// TIA Portal V20 export
FUNCTION_BLOCK "OP1"   // FB50, LAD
{ S7_Optimized_Access := 'TRUE' }
// stored: AutoNumber false, MemoryReserve 100, SetENOAutomatically false
   VAR DB_SPECIFIC
      CONTROL_MAN : Struct
         kar_work : Bool;
         kar_home : Bool;
         zarazka_work : Bool;
         zarazka_home : Bool;
         B4 : Bool;
         B5 : Bool;
         B6 : Bool;
         B7 : Bool;
         B8 : Bool;
         B9 : Bool;
         odfuk_1 : Bool;
         odfuk_2 : Bool;
         B12 : Bool;
         B13 : Bool;
         B14 : Bool;
         B15 : Bool;
         B16 : Bool;
         B17 : Bool;
         B18 : Bool;
         B19 : Bool;
         B20 : Bool;
         B21 : Bool;
         B22 : Bool;
         B23 : Bool;
         B24 : Bool;
         B25 : Bool;
         B26 : Bool;
         B27 : Bool;
         B28 : Bool;
         B29 : Bool;
         B30 : Bool;
         B31 : Bool;
      END_STRUCT;
      CONTROL_AUTOMAT : Struct
         KAR_WORK : Bool;
         KAR_HOME : Bool;
         ZARAZKA_WORK : Bool;
         ZARAZKA_HOME : Bool;
         B4 : Bool;
         B5 : Bool;
         B6 : Bool;
         B7 : Bool;
         B8 : Bool;
         B9 : Bool;
         odfuk_1 : Bool;
         odfuk_2 : Bool;
         B12 : Bool;
         B13 : Bool;
         B14 : Bool;
         B15 : Bool;
         B16 : Bool;
         B17 : Bool;
         B18 : Bool;
         B19 : Bool;
         B20 : Bool;
         B21 : Bool;
         B22 : Bool;
         B23 : Bool;
         B24 : Bool;
         B25 : Bool;
         B26 : Bool;
         B27 : Bool;
         B28 : Bool;
         B29 : Bool;
         B30 : Bool;
         B31 : Bool;
      END_STRUCT;
      SENSORS : Struct
         prechod_1 : Bool;
         prechod_1_neg : Bool;
         kontrola : Bool;
         kontrola_neg : Bool;
         prechod_2 : Bool;
         Prechod_2_neg : Bool;
         Pozice_vyrazovace : Bool;
         Pozice_vyrazovace_neg : Bool;
         Pozice_pistu : Bool;   // KARUSEL JE NATOČEN PŘÍPRAVKEM A K BRÁNĚ
         Pozice_pistu_neg : Bool;
         s10 : Bool;
         s11 : Bool;
         s12 : Bool;
         s13 : Bool;
         s14 : Bool;
         s15 : Bool;
         s16 : Bool;
         s17 : Bool;
         s18 : Bool;
         s19 : Bool;
         s20 : Bool;
         s21 : Bool;
         s22 : Bool;
         s23 : Bool;
         s24 : Bool;
         s25 : Bool;
         s26 : Bool;
         s27 : Bool;
         s28 : Bool;
         s29 : Bool;
         s30 : Bool;
         s31 : Bool;
      END_STRUCT;
      SENSORS_1 : Struct
         S0 : Bool;
         S1 : Bool;
         S2 : Bool;
         S3 : Bool;
         S4 : Bool;
         S5 : Bool;
         S6 : Bool;
         S7 : Bool;
         S8 : Bool;
         S9 : Bool;
         SESTAVA_NENI_OTOCENA : Bool;
         SESTAVA_JE_OTOCENA : Bool;
         S12 : Bool;
         S13 : Bool;
         S14 : Bool;
         S15 : Bool;
         S16 : Bool;
         S17 : Bool;
         S18 : Bool;
         S19 : Bool;
         S20 : Bool;
         S21 : Bool;
         S22 : Bool;
         S23 : Bool;
         S24 : Bool;
         S25 : Bool;
         S26 : Bool;
         S27 : Bool;
         S28 : Bool;
         S29 : Bool;
         S30 : Bool;
         l_3_neg : Bool;
      END_STRUCT;
   END_VAR
   VAR
      S_0 : "SENSOR";
      S_1 : "SENSOR";
      S_2 { S7_SetPoint := 'True'} : "SENSOR";
      S_3 { S7_SetPoint := 'True'} : "SENSOR";
      S_4 { S7_SetPoint := 'True'} : "SENSOR";
      S_5 { S7_SetPoint := 'True'} : "SENSOR";
      S_6 { S7_SetPoint := 'True'} : "SENSOR";
      M_karusel : "MOTOR_CONTROL_BLOCK";
      M_zarazka { S7_SetPoint := 'True'} : "MOTOR_CONTROL_BLOCK";
      M_CLONA { S7_SetPoint := 'True'} : "MOTOR_CONTROL_BLOCK";
   END_VAR
   VAR DB_SPECIFIC
      SQCR { S7_SetPoint := 'True'} : Int;
   END_VAR
   VAR
      hmi_sqcr : Int;
   END_VAR
   VAR DB_SPECIFIC
      TRIG : Struct
         inicial_ok_op : Bool;
         DSSAD : Bool;
         INICIALIZACE_PROBEHLA : Bool;
         trig_dil : Bool;
         p_trig_control_tcon : Bool;
         T6 : Bool;
         SPUST_OP_4 : Bool;
         vlez_do_zavory_pri_rotaci : Bool;
         START_INICIAL_OP2 : Bool;
         START_INICIAL_OP3 : Bool;
         spust_odsavani : Bool;
         VYPRAZNI_OK_OP_2_A : Bool;
         VYPRAZNI_NOK_OP_2_A : Bool;
         VYPRAZDNI_OK_OP_3_B : Bool;
         VYPRAZDNI_NOK_OP_3_B : Bool;
         RESET_NCODER : Bool;
         op_1_ready : Bool;
      END_STRUCT;
      MEMOR : Struct
         n_trig_vypnuti : Bool;
         M1 : Bool;
         M2 : Bool;
         M3 : Bool;
         M4 : Bool;
         p_trig_odavacka : Bool;
         M6 : Bool;
         M7 : Bool;
         M8 : Bool;
         M9 : Bool;
         M10 : Bool;
         M11 : Bool;
         RESET_ERROR : Bool;
         vyrazeni_pamet : Bool;
         M14 : Bool;
         M15 : Bool;
         SETOVANI_START : Bool;
         M17 : Bool;
         p_trig_pamet_1 : Bool;
         p_trig_pamet_2 : Bool;
         p_trig_pamet_3 : Bool;
         p_trig_pamet_4 : Bool;
         p_trig_pamet_5 : Bool;
         p_trig_pamet_6 : Bool;
         p_trig_pamet_7 : Bool;
         p_trig_pamet_8 : Bool;
         p_trig_pamet_9 : Bool;
         p_trig_pamet_10 : Bool;
         p_trig_vyrad : Bool;
         p_Trig_cisteni_pozice : Bool;
         p_trig_citac : Bool;
         N_TRIG_SAFETY : Bool;
         P_TRIG_RESET_POZICE : Bool;
         M33 : Bool;
         start_caklu : Bool;
         M35 : Bool;
         M36 : Bool;
         M37 : Bool;
         M38 : Bool;
         M39 : Bool;
         ALARM_GLOBAL : Bool;
         M41 : Bool;
         M42 : Bool;
         M43 : Bool;
         M44 : Bool;
         M45 : Bool;
         M46 : Bool;
         M47 : Bool;
         M48 : Bool;
         M49 : Bool;
         wrong_p_trig : Bool;
         alarm_p_trig : Bool;
         M52 : Bool;
         M53 : Bool;
         M54 : Bool;
         M55 : Bool;
         M56 : Bool;
         M57 : Bool;
         M58 : Bool;
         M59 : Bool;
         M60 : Bool;
         M61 : Bool;
         M62 : Bool;
         M63 : Bool;
      END_STRUCT;
      "TIMER" : Struct
         TIMER_0 : IEC_TIMER;
         TIMER_VACUUM_CLEANER : IEC_TIMER;
         TIMER_DELAY_RESET_EXECUTE : IEC_TIMER;
         TIMER_3 : IEC_TIMER;
         TIMER_4 : IEC_TIMER;
         air : IEC_TIMER;
         TIMER_6 : IEC_TIMER;
         TIMER_7 : IEC_TIMER;
      END_STRUCT;
      HMI : Struct
         povoleni_volby_receptu : Bool;
         "svetlo_on/off" : Bool;
         ALARM_VIDITELNOST : Bool;
         hmi_3 : Bool;
         hmi_4 : Bool;
         reset_fronty : Bool;
         hmi_6 : Bool;
         hmi_7 : Bool;
         hmi_8 : Bool;
         hmi_9 : Bool;
         hmi_10 : Bool;
         hmi_11 : Bool;
         hmi_12 : Bool;
         hmi_13 : Bool;
         hmi_14 : Bool;
         hmi_15 : Bool;
      END_STRUCT;
   END_VAR
   VAR
      STRING_0 : String[1];
      array_chyb_ctec : Array[1..16] of Bool;
      zpracovani_dat { ExternalAccessible := 'False'; ExternalVisible := 'False'; ExternalWritable := 'False'} : Array[1..1] of Struct
         prenaseny_text : String[100];
         balik_den : Int;
         vyrazeni : Bool;
      END_STRUCT;
   END_VAR
   VAR DB_SPECIFIC
      aktual_kusy : Int;
   END_VAR
   VAR
      i : Int;
      q : Int;
      pocet_znaku_string_kamera : Int;
      ocekavany_text : String[100];
      format_etiketa_ok : Bool;
      Kamera : Struct
         s2_pamet : Bool;
         s2_nabeh : Bool;
         sber_aktivni : Bool;
         prijato_etiketa : Bool;
         prijato_folie_l : Bool;
         prijato_folie_p : Bool;
         ok_etiketa : Bool;
         ok_folie_l : Bool;
         ok_folie_p : Bool;
         vyradit : Bool;
         fronta_plna : Bool;   // alarm
         bypass_ocr : Bool := True;   // dočasně, dokud není doladěné OCR
         last_id_etiketa : Word;
         last_id_folie_l : Word;
         last_id_folie_p : Word;
         balik_den : Int;
         idx : Int;
         pocet : Int;
         text_etiketa : String[100];
         timeout_sberu : Time :=  T#1S;
         kontrola_tridirny : Bool := true;   // HMI: kontrola kódu třídírny zapnuta
         tridirna_ok : Bool;   // výsledek kontroly posledního plata (pro online diagnostiku)
      END_STRUCT;
      Vyrazeni : Struct
         s4_pamet : Bool;
         s4_nabeh : Bool;
         aktivni : Bool;
         vyradit : Bool;
         chyba_bez_dat : Bool;   // alarm: plato u vyřazovače bez záznamu
         chyba_pist : Bool;   // alarm: píst nevyjel / nebyl v home
         max_puls : Time := T#200MS;
         vyrazovac_pripojen : Bool := true;   // TRUE až bude signál od dodavatele
         alarm_nok_balik : Bool;   // NOK plato prošlo bez vyřazení
         posledni_nok_balik : Int;   // číslo plata pro obsluhu / HMI
         posledni_nok_text : String[100];   // co přečetla kamera
         pocet_nok : DInt;   // počítadlo NOK plat
         pocet_bez_dat : DInt;
         majak_tp : TP_TIME;   // prodlouzeni blikani majaku pri vzrazenii
         majak { S7_SetPoint := 'True'} : Bool;
      END_STRUCT;
      Kam_Etiketa_Job : Struct
         krok : Int;   // 0 klid, 10 odeslat, 20 čekat, 30 ukončit handshake
         pozadovany : Int;   // job z receptury (PRG_CAM_etiketa)
         odesli_pamet : Bool;   // hrana ODESLI_dATA
         aktivni : Bool;   // probíhá načítání jobu → blokovat triggery
         chyba : Bool;   // alarm: job se nepodařilo načíst
         chyba_kod : Word;   // CommandResultCode při chybě
         nesouhlasi : Bool;   // alarm: job v kameře ≠ job z receptury
         timeout : Time := T#10S;   // max. doba načítání jobu
      END_STRUCT;
      Test_tp_ka12 : TP_TIME;
   END_VAR
   VAR_TEMP
      DATA : Array[0..255] of Char;
      ARRAY_NULL : Array[1..8] of Bool;
      array_null_fronta : Array[1..1] of Struct
         prenaseny_text : String[100];
         balik_den : Int;
         vyrazeni : Bool;
      END_STRUCT;
      "char" : Array[0..0] of Char;
      "string" : String;
      cas : DTL;
      ret : Int;
   END_VAR
   VAR CONSTANT
      STEP_0 : Int := 0;
      step_2 : Int := 2;
      STEP_4 : Int := 4;
      STEP_5_HOME : Int := 5;
      STEP_7 : Int := 7;
      STEP_10 : Int := 10;
      STEP_15 : Int := 15;
      STEP_20 : Int := 20;
      STEP_23 : Int := 23;
      STEP_25 : Int := 25;
      STEP_27 : Int := 27;
      STEP_30 : Int := 30;
      STEP_35 : Int := 35;
      STEP_37 : Int := 37;
      STEP_40 : Int := 40;
      STEP_45 : Int := 45;
      STEP_50 : Int := 50;
      STEP_55 : Int := 55;
      STEP_60 : Int := 60;
      STEP_65 : Int := 65;
      STEP_70 : Int := 70;
      STEP_75 : Int := 75;
      STEP_80 : Int := 80;
      STEP_83 : Int := 83;
      STEP_85 : Int := 85;
      STEP_90 : Int := 90;
      STEP_95 : Int := 95;
      STEP_100 : Int := 100;
      STEP_105 : Int := 105;
      STEP_110 : Int := 110;
      STEP_113 : Int := 113;
      STEP_115 : Int := 115;
      STEP_120 : Int := 120;
      STEP_125 : Int := 125;
      STEP_130 : Int := 130;
      STEP_135 : Int := 135;
      STEP_140 : Int := 140;
      STEP_145 : Int := 145;
      STEP_150 : Int := 150;
      STEP_155 : Int := 155;
      STEP_1000 : Int := 1000;
      STEP_1001 : Int := 1001;
      STEP_1002 : Int := 1002;
      STEP_1003 : Int := 1003;
      STEP_1004 : Int := 1004;
      STEP_1005 : Int := 1005;
      STEP_1010 : Int := 1010;
      STEP_1015 : Int := 1015;
      STEP_1020 : Int := 1020;
      STEP_1025 : Int := 1025;
      STEP_3000 : Int := 3000;
      STEP_3005 : Int := 3005;
      STEP_3010 : Int := 3010;
      STEP_3015 : Int := 3015;
      STEP_3020 : Int := 3020;
      STEP_2000 : Int := 2000;
      string_null : String;
      char_null : Char;
      text_kartacek : String := 'Kartacek';
      string_kar_A : String := 'A';
      string_kar_B : String := 'B';
      KOD_TRIDIRNY : String := 'CZ32880102';
   END_VAR
   VAR_TEMP   // added for the SCL form of the ladder/FBD networks
      _w1 : Bool;
      _w2 : Bool;
      _w3 : Bool;
   END_VAR
BEGIN

REGION Network 1: manuali ovladani reset
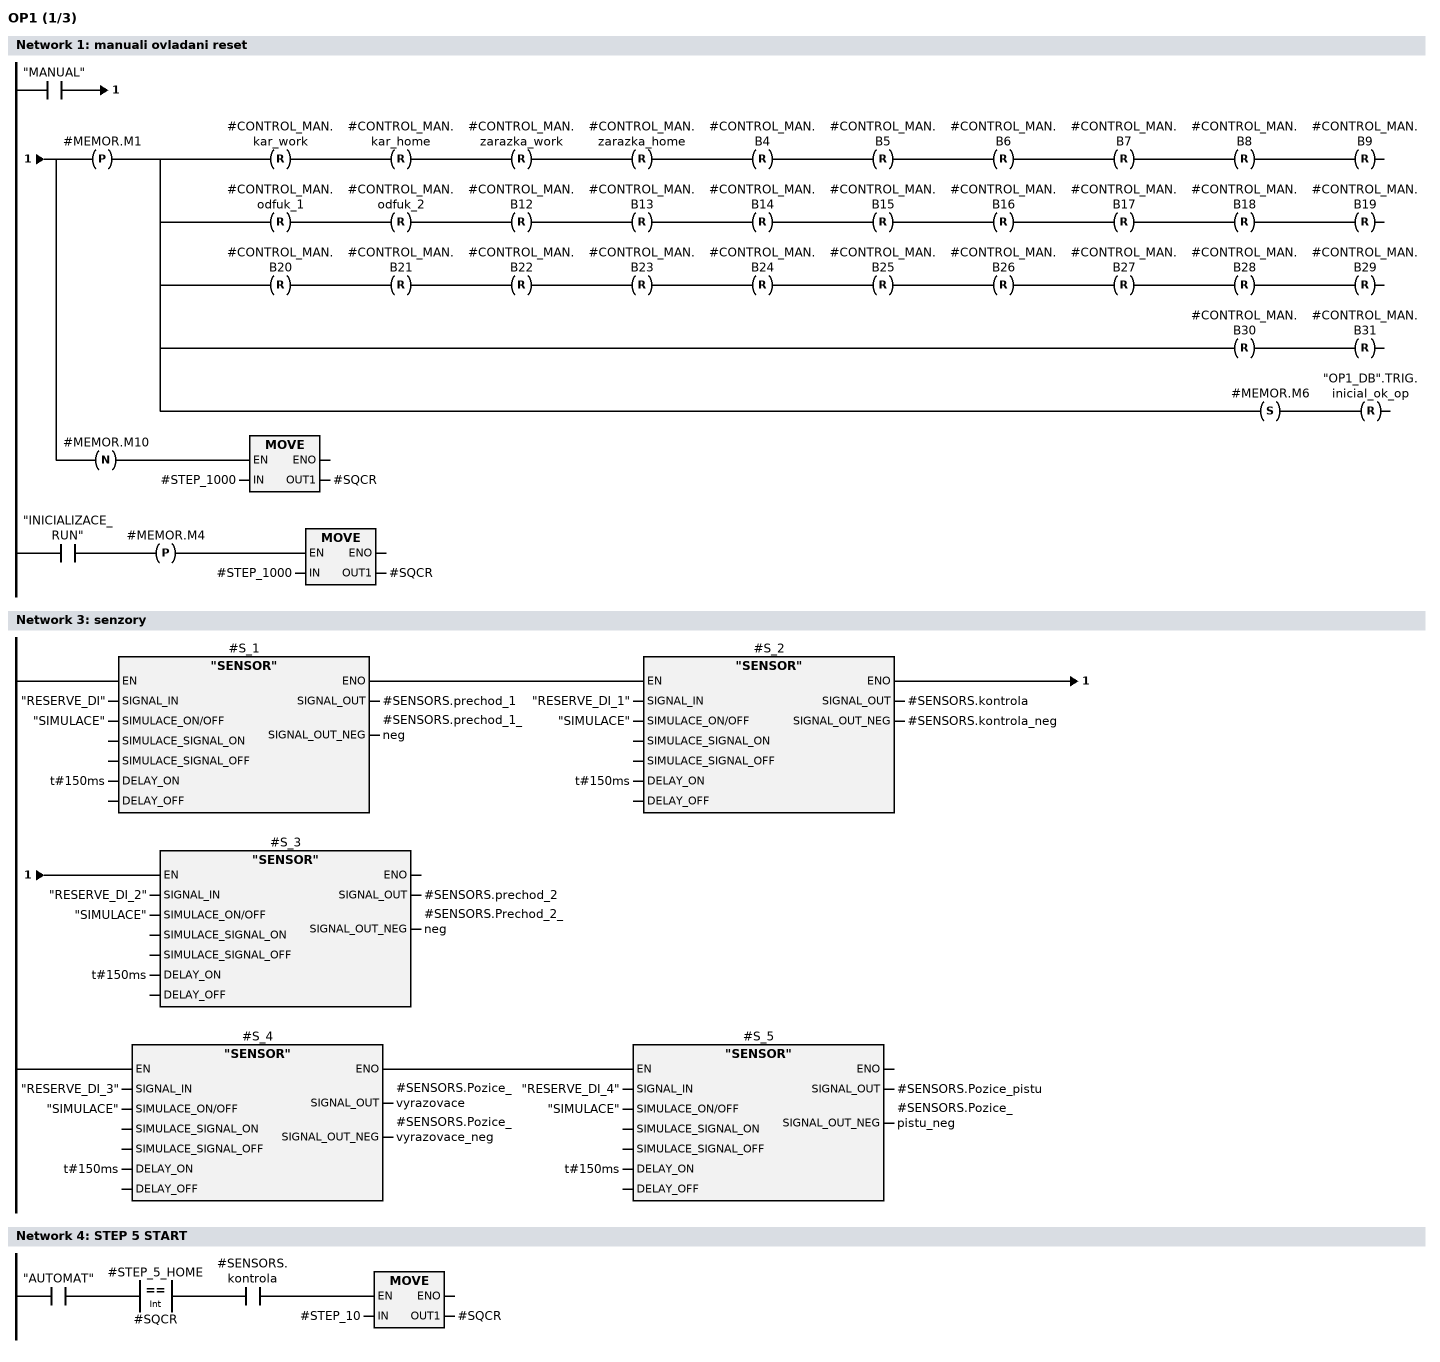
   RUNG wire#powerrail
      Contact( "MANUAL" )
      wire#w1
      P_Trig( #MEMOR.M1 )
      wire#w2
      R_Coil( #CONTROL_MAN.kar_work )
      R_Coil( #CONTROL_MAN.kar_home )
      R_Coil( #CONTROL_MAN.zarazka_work )
      R_Coil( #CONTROL_MAN.zarazka_home )
      R_Coil( #CONTROL_MAN.B4 )
      R_Coil( #CONTROL_MAN.B5 )
      R_Coil( #CONTROL_MAN.B6 )
      R_Coil( #CONTROL_MAN.B7 )
      R_Coil( #CONTROL_MAN.B8 )
      R_Coil( #CONTROL_MAN.B9 )
   END_RUNG
   RUNG wire#w2
      R_Coil( #CONTROL_MAN.odfuk_1 )
      R_Coil( #CONTROL_MAN.odfuk_2 )
      R_Coil( #CONTROL_MAN.B12 )
      R_Coil( #CONTROL_MAN.B13 )
      R_Coil( #CONTROL_MAN.B14 )
      R_Coil( #CONTROL_MAN.B15 )
      R_Coil( #CONTROL_MAN.B16 )
      R_Coil( #CONTROL_MAN.B17 )
      R_Coil( #CONTROL_MAN.B18 )
      R_Coil( #CONTROL_MAN.B19 )
   END_RUNG
   RUNG wire#w2
      R_Coil( #CONTROL_MAN.B20 )
      R_Coil( #CONTROL_MAN.B21 )
      R_Coil( #CONTROL_MAN.B22 )
      R_Coil( #CONTROL_MAN.B23 )
      R_Coil( #CONTROL_MAN.B24 )
      R_Coil( #CONTROL_MAN.B25 )
      R_Coil( #CONTROL_MAN.B26 )
      R_Coil( #CONTROL_MAN.B27 )
      R_Coil( #CONTROL_MAN.B28 )
      R_Coil( #CONTROL_MAN.B29 )
   END_RUNG
   RUNG wire#w2
      R_Coil( #CONTROL_MAN.B30 )
      R_Coil( #CONTROL_MAN.B31 )
   END_RUNG
   RUNG wire#w2
      S_Coil( #MEMOR.M6 )
      R_Coil( "OP1_DB".TRIG.inicial_ok_op )
   END_RUNG
   RUNG wire#w1
      N_Trig( #MEMOR.M10 )
      Move(in := #STEP_1000, out1 => #SQCR)
   END_RUNG
   RUNG wire#powerrail
      Contact( "INICIALIZACE_RUN" )
      P_Trig( #MEMOR.M4 )
      Move(in := #STEP_1000, out1 => #SQCR)
   END_RUNG
   // the same network as SCL:
   #_w1 := "MANUAL" AND NOT #MEMOR.M1;   // rising edge
   #MEMOR.M1 := "MANUAL";
   IF #_w1 THEN
       #CONTROL_MAN.kar_work := FALSE;
       #CONTROL_MAN.kar_home := FALSE;
       #CONTROL_MAN.zarazka_work := FALSE;
       #CONTROL_MAN.zarazka_home := FALSE;
       #CONTROL_MAN.B4 := FALSE;
       #CONTROL_MAN.B5 := FALSE;
       #CONTROL_MAN.B6 := FALSE;
       #CONTROL_MAN.B7 := FALSE;
       #CONTROL_MAN.B8 := FALSE;
       #CONTROL_MAN.B9 := FALSE;
       #CONTROL_MAN.odfuk_1 := FALSE;
       #CONTROL_MAN.odfuk_2 := FALSE;
       #CONTROL_MAN.B12 := FALSE;
       #CONTROL_MAN.B13 := FALSE;
       #CONTROL_MAN.B14 := FALSE;
       #CONTROL_MAN.B15 := FALSE;
       #CONTROL_MAN.B16 := FALSE;
       #CONTROL_MAN.B17 := FALSE;
       #CONTROL_MAN.B18 := FALSE;
       #CONTROL_MAN.B19 := FALSE;
       #CONTROL_MAN.B20 := FALSE;
       #CONTROL_MAN.B21 := FALSE;
       #CONTROL_MAN.B22 := FALSE;
       #CONTROL_MAN.B23 := FALSE;
       #CONTROL_MAN.B24 := FALSE;
       #CONTROL_MAN.B25 := FALSE;
       #CONTROL_MAN.B26 := FALSE;
       #CONTROL_MAN.B27 := FALSE;
       #CONTROL_MAN.B28 := FALSE;
       #CONTROL_MAN.B29 := FALSE;
       #CONTROL_MAN.B30 := FALSE;
       #CONTROL_MAN.B31 := FALSE;
       #MEMOR.M6 := TRUE;
       "OP1_DB".TRIG.inicial_ok_op := FALSE;
   END_IF;
   #_w2 := NOT "MANUAL" AND #MEMOR.M10;   // falling edge
   #MEMOR.M10 := "MANUAL";
   IF #_w2 THEN #SQCR := #STEP_1000; END_IF;
   #_w3 := "INICIALIZACE_RUN" AND NOT #MEMOR.M4;   // rising edge
   #MEMOR.M4 := "INICIALIZACE_RUN";
   IF #_w3 THEN #SQCR := #STEP_1000; END_IF;
END_REGION

REGION Network 2: alarmy
END_REGION

REGION Network 3: senzory
   RUNG wire#powerrail
      #S_1(SIGNAL_IN := "RESERVE_DI", "SIMULACE_ON/OFF" := "SIMULACE", SIMULACE_SIGNAL_ON :=, SIMULACE_SIGNAL_OFF :=, DELAY_ON := t#150ms, DELAY_OFF :=, SIGNAL_OUT => #SENSORS.prechod_1, SIGNAL_OUT_NEG => #SENSORS.prechod_1_neg)
      #S_2(SIGNAL_IN := "RESERVE_DI_1", "SIMULACE_ON/OFF" := "SIMULACE", SIMULACE_SIGNAL_ON :=, SIMULACE_SIGNAL_OFF :=, DELAY_ON := t#150ms, DELAY_OFF :=, SIGNAL_OUT => #SENSORS.kontrola, SIGNAL_OUT_NEG => #SENSORS.kontrola_neg)
      #S_3(SIGNAL_IN := "RESERVE_DI_2", "SIMULACE_ON/OFF" := "SIMULACE", SIMULACE_SIGNAL_ON :=, SIMULACE_SIGNAL_OFF :=, DELAY_ON := t#150ms, DELAY_OFF :=, SIGNAL_OUT => #SENSORS.prechod_2, SIGNAL_OUT_NEG => #SENSORS.Prechod_2_neg)
   END_RUNG
   RUNG wire#powerrail
      #S_4(SIGNAL_IN := "RESERVE_DI_3", "SIMULACE_ON/OFF" := "SIMULACE", SIMULACE_SIGNAL_ON :=, SIMULACE_SIGNAL_OFF :=, DELAY_ON := t#150ms, DELAY_OFF :=, SIGNAL_OUT => #SENSORS.Pozice_vyrazovace, SIGNAL_OUT_NEG => #SENSORS.Pozice_vyrazovace_neg)
      #S_5(SIGNAL_IN := "RESERVE_DI_4", "SIMULACE_ON/OFF" := "SIMULACE", SIMULACE_SIGNAL_ON :=, SIMULACE_SIGNAL_OFF :=, DELAY_ON := t#150ms, DELAY_OFF :=, SIGNAL_OUT => #SENSORS.Pozice_pistu, SIGNAL_OUT_NEG => #SENSORS.Pozice_pistu_neg)
   END_RUNG
   // the same network as SCL:
   #S_1(SIGNAL_IN := "RESERVE_DI",   // "SENSOR"
        "SIMULACE_ON/OFF" := "SIMULACE",
        DELAY_ON := t#150ms,
        SIGNAL_OUT => #SENSORS.prechod_1,
        SIGNAL_OUT_NEG => #SENSORS.prechod_1_neg,
        ENO => #_w1);
   #S_2(EN := #_w1,   // "SENSOR"
        SIGNAL_IN := "RESERVE_DI_1",
        "SIMULACE_ON/OFF" := "SIMULACE",
        DELAY_ON := t#150ms,
        SIGNAL_OUT => #SENSORS.kontrola,
        SIGNAL_OUT_NEG => #SENSORS.kontrola_neg,
        ENO => #_w2);
   IF #_w2 THEN
       #S_3(SIGNAL_IN := "RESERVE_DI_2",   // "SENSOR"
            "SIMULACE_ON/OFF" := "SIMULACE",
            DELAY_ON := t#150ms,
            SIGNAL_OUT => #SENSORS.prechod_2,
            SIGNAL_OUT_NEG => #SENSORS.Prechod_2_neg);
   END_IF;
   #S_4(SIGNAL_IN := "RESERVE_DI_3",   // "SENSOR"
        "SIMULACE_ON/OFF" := "SIMULACE",
        DELAY_ON := t#150ms,
        SIGNAL_OUT => #SENSORS.Pozice_vyrazovace,
        SIGNAL_OUT_NEG => #SENSORS.Pozice_vyrazovace_neg,
        ENO => #_w3);
   IF #_w3 THEN
       #S_5(SIGNAL_IN := "RESERVE_DI_4",   // "SENSOR"
            "SIMULACE_ON/OFF" := "SIMULACE",
            DELAY_ON := t#150ms,
            SIGNAL_OUT => #SENSORS.Pozice_pistu,
            SIGNAL_OUT_NEG => #SENSORS.Pozice_pistu_neg);
   END_IF;
END_REGION

REGION Network 4: STEP 5 START
   RUNG wire#powerrail
      Contact( "AUTOMAT" )
      { S7_Templates := "SrcType := Int" } EQ_Contact(in1 := #STEP_5_HOME, in2 := #SQCR)
      Contact( #SENSORS.kontrola )
      Move(in := #STEP_10, out1 => #SQCR)
   END_RUNG
   // the same network as SCL:
   IF "AUTOMAT" AND (#STEP_5_HOME = #SQCR) AND #SENSORS.kontrola THEN #SQCR := #STEP_10; END_IF;
END_REGION

REGION Network 5: STEP 10
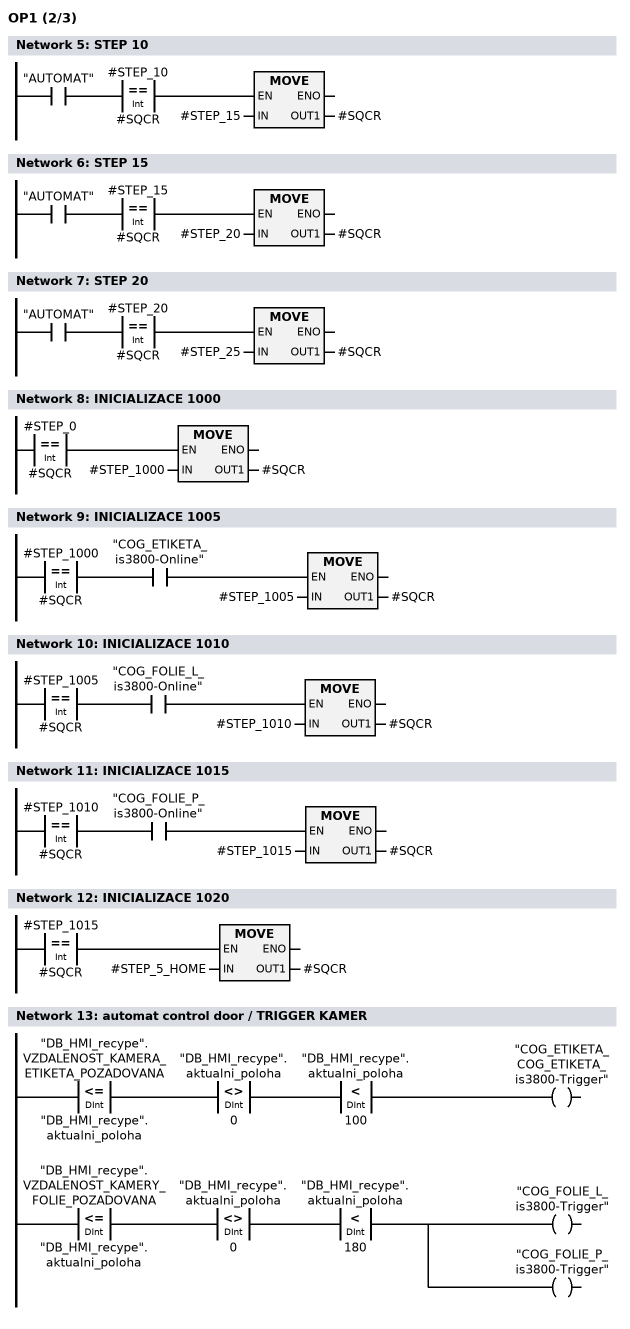
   RUNG wire#powerrail
      Contact( "AUTOMAT" )
      { S7_Templates := "SrcType := Int" } EQ_Contact(in1 := #STEP_10, in2 := #SQCR)
      Move(in := #STEP_15, out1 => #SQCR)
   END_RUNG
   // the same network as SCL:
   IF "AUTOMAT" AND (#STEP_10 = #SQCR) THEN #SQCR := #STEP_15; END_IF;
END_REGION

REGION Network 6: STEP 15
   RUNG wire#powerrail
      Contact( "AUTOMAT" )
      { S7_Templates := "SrcType := Int" } EQ_Contact(in1 := #STEP_15, in2 := #SQCR)
      Move(in := #STEP_20, out1 => #SQCR)
   END_RUNG
   // the same network as SCL:
   IF "AUTOMAT" AND (#STEP_15 = #SQCR) THEN #SQCR := #STEP_20; END_IF;
END_REGION

REGION Network 7: STEP 20
   RUNG wire#powerrail
      Contact( "AUTOMAT" )
      { S7_Templates := "SrcType := Int" } EQ_Contact(in1 := #STEP_20, in2 := #SQCR)
      Move(in := #STEP_25, out1 => #SQCR)
   END_RUNG
   // the same network as SCL:
   IF "AUTOMAT" AND (#STEP_20 = #SQCR) THEN #SQCR := #STEP_25; END_IF;
END_REGION

REGION Network 8: INICIALIZACE 1000
   RUNG wire#powerrail
      { S7_Templates := "SrcType := Int" } EQ_Contact(in1 := #STEP_0, in2 := #SQCR)
      Move(in := #STEP_1000, out1 => #SQCR)
   END_RUNG
   // the same network as SCL:
   IF #STEP_0 = #SQCR THEN #SQCR := #STEP_1000; END_IF;
END_REGION

REGION Network 9: INICIALIZACE 1005
   RUNG wire#powerrail
      { S7_Templates := "SrcType := Int" } EQ_Contact(in1 := #STEP_1000, in2 := #SQCR)
      Contact( "COG_ETIKETA_is3800-Online" )
      Move(in := #STEP_1005, out1 => #SQCR)
   END_RUNG
   // the same network as SCL:
   IF (#STEP_1000 = #SQCR) AND "COG_ETIKETA_is3800-Online" THEN #SQCR := #STEP_1005; END_IF;
END_REGION

REGION Network 10: INICIALIZACE 1010
   RUNG wire#powerrail
      { S7_Templates := "SrcType := Int" } EQ_Contact(in1 := #STEP_1005, in2 := #SQCR)
      Contact( "COG_FOLIE_L_is3800-Online" )
      Move(in := #STEP_1010, out1 => #SQCR)
   END_RUNG
   // the same network as SCL:
   IF (#STEP_1005 = #SQCR) AND "COG_FOLIE_L_is3800-Online" THEN #SQCR := #STEP_1010; END_IF;
END_REGION

REGION Network 11: INICIALIZACE 1015
   RUNG wire#powerrail
      { S7_Templates := "SrcType := Int" } EQ_Contact(in1 := #STEP_1010, in2 := #SQCR)
      Contact( "COG_FOLIE_P_is3800-Online" )
      Move(in := #STEP_1015, out1 => #SQCR)
   END_RUNG
   // the same network as SCL:
   IF (#STEP_1010 = #SQCR) AND "COG_FOLIE_P_is3800-Online" THEN #SQCR := #STEP_1015; END_IF;
END_REGION

REGION Network 12: INICIALIZACE 1020
   RUNG wire#powerrail
      { S7_Templates := "SrcType := Int" } EQ_Contact(in1 := #STEP_1015, in2 := #SQCR)
      Move(in := #STEP_5_HOME, out1 => #SQCR)
   END_RUNG
   // the same network as SCL:
   IF #STEP_1015 = #SQCR THEN #SQCR := #STEP_5_HOME; END_IF;
END_REGION

REGION Network 13: automat control door / TRIGGER KAMER
   RUNG wire#powerrail
      { S7_Templates := "SrcType := DInt" } LE_Contact(in1 := "DB_HMI_recype".VZDALENOST_KAMERA_ETIKETA_POZADOVANA, in2 := "DB_HMI_recype".aktualni_poloha)
      { S7_Templates := "SrcType := DInt" } NE_Contact(in1 := "DB_HMI_recype".aktualni_poloha, in2 := 0)
      { S7_Templates := "SrcType := DInt" } LT_Contact(in1 := "DB_HMI_recype".aktualni_poloha, in2 := 100)
      Coil( "COG_ETIKETA_COG_ETIKETA_is3800-Trigger" )
   END_RUNG
   RUNG wire#powerrail
      { S7_Templates := "SrcType := DInt" } LE_Contact(in1 := "DB_HMI_recype".VZDALENOST_KAMERY_FOLIE_POZADOVANA, in2 := "DB_HMI_recype".aktualni_poloha)
      { S7_Templates := "SrcType := DInt" } NE_Contact(in1 := "DB_HMI_recype".aktualni_poloha, in2 := 0)
      { S7_Templates := "SrcType := DInt" } LT_Contact(in1 := "DB_HMI_recype".aktualni_poloha, in2 := 180)
      wire#w1
      Coil( "COG_FOLIE_L_is3800-Trigger" )
   END_RUNG
   RUNG wire#w1
      Coil( "COG_FOLIE_P_is3800-Trigger" )
   END_RUNG
   // the same network as SCL:
   "COG_ETIKETA_COG_ETIKETA_is3800-Trigger" := ("DB_HMI_recype".VZDALENOST_KAMERA_ETIKETA_POZADOVANA <= "DB_HMI_recype".aktualni_poloha) AND ("DB_HMI_recype".aktualni_poloha <> 0) AND ("DB_HMI_recype".aktualni_poloha < 100);
   "COG_FOLIE_L_is3800-Trigger" := ("DB_HMI_recype".VZDALENOST_KAMERY_FOLIE_POZADOVANA <= "DB_HMI_recype".aktualni_poloha) AND ("DB_HMI_recype".aktualni_poloha <> 0) AND ("DB_HMI_recype".aktualni_poloha < 180);
   "COG_FOLIE_P_is3800-Trigger" := "COG_FOLIE_L_is3800-Trigger";
END_REGION

REGION Network 14: TRIGGER SVETEL
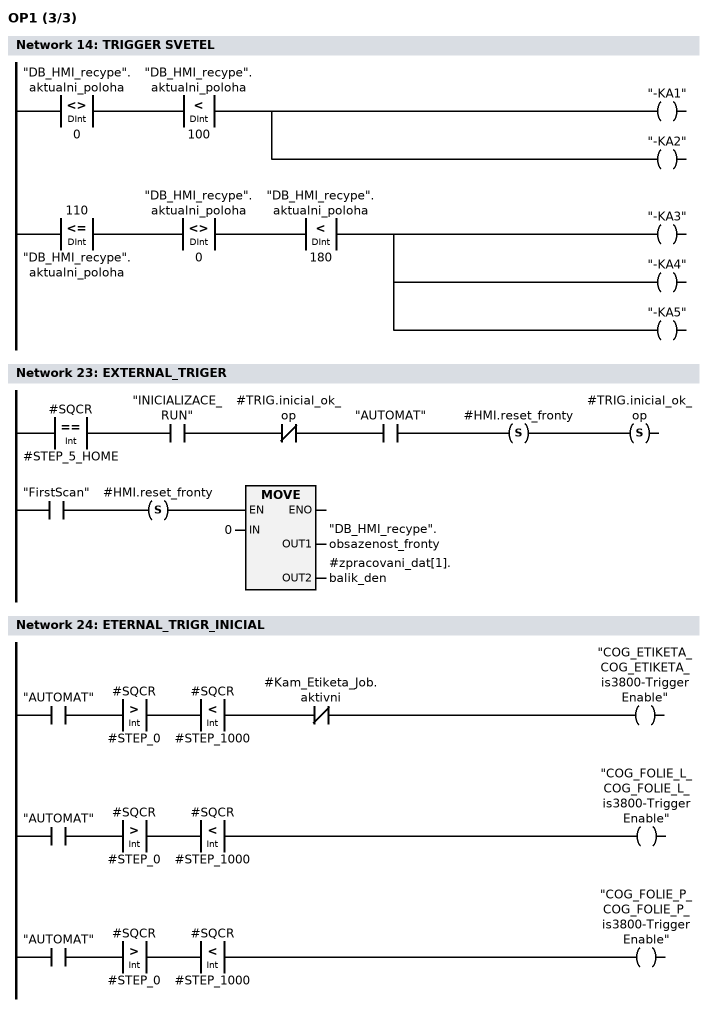
   RUNG wire#powerrail
      { S7_Templates := "SrcType := DInt" } NE_Contact(in1 := "DB_HMI_recype".aktualni_poloha, in2 := 0)
      { S7_Templates := "SrcType := DInt" } LT_Contact(in1 := "DB_HMI_recype".aktualni_poloha, in2 := 100)
      wire#w1
      Coil( "-KA1" )
   END_RUNG
   RUNG wire#w1
      Coil( "-KA2" )
   END_RUNG
   RUNG wire#powerrail
      { S7_Templates := "SrcType := DInt" } LE_Contact(in1 := 110, in2 := "DB_HMI_recype".aktualni_poloha)
      { S7_Templates := "SrcType := DInt" } NE_Contact(in1 := "DB_HMI_recype".aktualni_poloha, in2 := 0)
      { S7_Templates := "SrcType := DInt" } LT_Contact(in1 := "DB_HMI_recype".aktualni_poloha, in2 := 180)
      wire#w2
      Coil( "-KA3" )
   END_RUNG
   RUNG wire#w2
      Coil( "-KA4" )
   END_RUNG
   RUNG wire#w2
      Coil( "-KA5" )
   END_RUNG
   // the same network as SCL:
   "-KA1" := ("DB_HMI_recype".aktualni_poloha <> 0) AND ("DB_HMI_recype".aktualni_poloha < 100);
   "-KA2" := "-KA1";
   "-KA3" := (110 <= "DB_HMI_recype".aktualni_poloha) AND ("DB_HMI_recype".aktualni_poloha <> 0) AND ("DB_HMI_recype".aktualni_poloha < 180);
   "-KA4" := "-KA3";
   "-KA5" := "-KA3";
END_REGION

REGION Network 15 (SCL): TRIGGER MANUAL
   "iDB_CamManual"(xManEtiketa:="DB_Manual".xManEtiketa,
                   xManFolie:="DB_Manual".xManFolie);
END_REGION

REGION Network 16 (SCL): automat control data
   // Smyčka projde 104 bajtů (od 0 do 103)
   FOR #i := 0 TO 103 DO
       // PEEK čte přímo z paměti vstupů (16#81 = Periferní vstupy / Vstupy)
       // area 16#81 čte adresy %IB
       "DB_data_ctena".array_of_char[#i] := PEEK_BYTE(area := 16#81,
                                                       dbNumber := 0,
                                                       byteOffset := 76 + #i);
   END_FOR;

   // slozit text z prijatych znaku az po prvni $00
   "DB_data_ctena".upraveny := '';
   FOR #i := 0 TO 103 DO
       IF "DB_data_ctena".array_of_char[#i] = '$00' THEN
           EXIT;
       END_IF;
       "DB_data_ctena".upraveny := CONCAT(IN1 := "DB_data_ctena".upraveny,
                                          IN2 := CHAR_TO_STRING("DB_data_ctena".array_of_char[#i]));
   END_FOR;
END_REGION

REGION Network 17: automat control odfuk
END_REGION

REGION Network 18 (SCL): VYŘAZENÍ
   #Vyrazeni.s4_nabeh := #SENSORS.Pozice_vyrazovace AND NOT #Vyrazeni.s4_pamet;
   #Vyrazeni.s4_pamet := #SENSORS.Pozice_vyrazovace;

   IF "CONTROL_LINE_DB".trig.reset_error_all THEN
       #Vyrazeni.chyba_bez_dat := FALSE;
       #Vyrazeni.chyba_pist := FALSE;
       #Vyrazeni.alarm_nok_balik := FALSE;
   END_IF;

   IF NOT "AUTOMAT" THEN
       #Vyrazeni.aktivni := FALSE;
       #TIMER.TIMER_7.TON(IN := FALSE,
                          PT := #Vyrazeni.max_puls);
   ELSE
       REGION Plato prijelo k vyrazovaci - vzdy spotrebovat fronta[1]
           IF #Vyrazeni.s4_nabeh THEN
               IF "DB_HMI_recype".fronta[1].prenaseny_text = '' THEN
                   #Vyrazeni.chyba_bez_dat := TRUE;    // plato bez zaznamu ve fronte
                   #Vyrazeni.pocet_bez_dat := #Vyrazeni.pocet_bez_dat + 1;
                   #Vyrazeni.vyradit := TRUE;
               ELSE
                   #Vyrazeni.vyradit := "DB_HMI_recype".fronta[1].vyrazeni;
               END_IF;

               IF #Vyrazeni.vyradit THEN
                   #Vyrazeni.pocet_nok := #Vyrazeni.pocet_nok + 1;
                   IF "DB_HMI_recype".fronta[1].prenaseny_text = '' THEN
                       #Vyrazeni.posledni_nok_text := 'BEZ ZAZNAMU';
                       #Vyrazeni.posledni_nok_balik := 0;
                   ELSE
                       #Vyrazeni.posledni_nok_text := "DB_HMI_recype".fronta[1].prenaseny_text;
                       #Vyrazeni.posledni_nok_balik := "DB_HMI_recype".fronta[1].balik_den;
                   END_IF;
               END_IF;

               "DB_HMI_recype".fronta[1].prenaseny_text := '';
               "DB_HMI_recype".fronta[1].balik_den := 0;
               "DB_HMI_recype".fronta[1].vyrazeni := FALSE;

               IF #Vyrazeni.vyradit THEN
                   IF #Vyrazeni.vyrazovac_pripojen AND "DB_HMI_recype".recipe.vyrazovac_on_off THEN
                       #Vyrazeni.aktivni := TRUE;
                   ELSE
                       #Vyrazeni.alarm_nok_balik := TRUE;
                   END_IF;
               END_IF;
           END_IF;
       END_REGION

       REGION Pulz na vyrazovac - pevna delka Vyr.max_puls (200 ms)
           #TIMER.TIMER_7.TON(IN := #Vyrazeni.aktivni,
                              PT := #Vyrazeni.max_puls);
           IF #TIMER.TIMER_7.Q THEN
               #Vyrazeni.aktivni := FALSE;
           END_IF;
       END_REGION
   END_IF;

   // vystup na vyrazovac + rucni test (DB_Manual.test_vyr drzi vystup, dokud je TRUE)
   "RESERVE_DQ_2" := (#Vyrazeni.aktivni AND #Vyrazeni.vyrazovac_pripojen) OR "DB_Manual".test_vyr;

   // majak: po kazdem vyrazeni blika 5 s
   #Vyrazeni.majak_tp(IN := #Vyrazeni.aktivni AND #Vyrazeni.vyrazovac_pripojen,
                      PT := T#3S);
   #Vyrazeni.majak := #Vyrazeni.majak_tp.Q;
END_REGION

REGION Network 19 (SCL): CONTROL BLOCK presun_fronty
   IF "AUTOMAT" = true THEN


       REGION fronta 1 z 2
           IF "DB_HMI_recype".fronta[1].prenaseny_text = '' AND "DB_HMI_recype".fronta[2].prenaseny_text <> '' THEN
               "DB_HMI_recype".fronta[1]:= "DB_HMI_recype".fronta[2];
               "DB_HMI_recype".fronta[2].prenaseny_text := '';
               "DB_HMI_recype".fronta[2].balik_den := 0;
               "DB_HMI_recype".fronta[2].vyrazeni := false;
           END_IF;
       END_REGION

       REGION fronta 2 z 3
           IF "DB_HMI_recype".fronta[2].prenaseny_text = '' AND "DB_HMI_recype".fronta[3].prenaseny_text <> '' THEN
               "DB_HMI_recype".fronta[2] := "DB_HMI_recype".fronta[3];
               "DB_HMI_recype".fronta[3].prenaseny_text := '';
               "DB_HMI_recype".fronta[3].balik_den := 0;
               "DB_HMI_recype".fronta[3].vyrazeni := false;
           END_IF;
       END_REGION

       REGION fronta 3 z 4
           IF "DB_HMI_recype".fronta[3].prenaseny_text = '' AND "DB_HMI_recype".fronta[4].prenaseny_text <> '' THEN
               "DB_HMI_recype".fronta[3] := "DB_HMI_recype".fronta[4];
               "DB_HMI_recype".fronta[4].prenaseny_text := '';
               "DB_HMI_recype".fronta[4].balik_den := 0;
               "DB_HMI_recype".fronta[4].vyrazeni := false;
           END_IF;
       END_REGION

       REGION fronta 4 z 5
           IF "DB_HMI_recype".fronta[4].prenaseny_text = '' AND "DB_HMI_recype".fronta[5].prenaseny_text <> '' THEN
               "DB_HMI_recype".fronta[4] := "DB_HMI_recype".fronta[5];
               "DB_HMI_recype".fronta[5].prenaseny_text := '';
               "DB_HMI_recype".fronta[5].balik_den := 0;
               "DB_HMI_recype".fronta[5].vyrazeni := false;
           END_IF;
       END_REGION



   END_IF;


   REGION mazání fronty operátorem - bude pak možnost i automaticky ?
   IF #HMI.reset_fronty = true THEN

       "DB_HMI_recype".fronta[1].prenaseny_text := '';
       "DB_HMI_recype".fronta[1].balik_den := 0;
       "DB_HMI_recype".fronta[1].vyrazeni := false;

       "DB_HMI_recype".fronta[2].prenaseny_text := '';
       "DB_HMI_recype".fronta[2].balik_den := 0;
       "DB_HMI_recype".fronta[2].vyrazeni := false;

       "DB_HMI_recype".fronta[3].prenaseny_text := '';
       "DB_HMI_recype".fronta[3].balik_den := 0;
       "DB_HMI_recype".fronta[3].vyrazeni := false;

       "DB_HMI_recype".fronta[4].prenaseny_text := '';
       "DB_HMI_recype".fronta[4].balik_den := 0;
       "DB_HMI_recype".fronta[4].vyrazeni := false;

       "DB_HMI_recype".fronta[5].prenaseny_text := '';
       "DB_HMI_recype".fronta[5].balik_den := 0;
       "DB_HMI_recype".fronta[5].vyrazeni := false;

       "DB_HMI_recype".obsazenost_fronty := 0;
       #HMI.reset_fronty := false;

   END_IF;
   END_REGION;
END_REGION

REGION Network 20 (SCL)
   // ===== DENNI RESET POCITADLA PLAT (o pulnoci, lokalni cas) =====
   #ret := RD_LOC_T(#cas);
   IF #cas.HOUR = 0 AND #cas.MINUTE = 0 AND #cas.SECOND = 0 THEN
       #zpracovani_dat[1].balik_den := 0;
   END_IF;
   #aktual_kusy := #zpracovani_dat[1].balik_den;
END_REGION

REGION Network 21 (SCL): SBĚR VÝSLEDKŮ A ZÁPIS DO FRONTY
   #Kamera.s2_nabeh := #SENSORS.kontrola AND NOT #Kamera.s2_pamet;
   #Kamera.s2_pamet := #SENSORS.kontrola;

   IF NOT "AUTOMAT" THEN
       #Kamera.sber_aktivni := FALSE;
       #Kamera.last_id_etiketa := "COG_ETIKETA_is3800-InspectionID";
       #Kamera.last_id_folie_l := "COG_FOLIE_L_is3800-InspectionID";
       #Kamera.last_id_folie_p := "COG_FOLIE_P_is3800-InspectionID";
       #TIMER.TIMER_6.TON(IN := FALSE,
                          PT := #Kamera.timeout_sberu);
   ELSE
       REGION Prijem vysledku (zmena InspectionID = dokoncena inspekce)
           IF "COG_ETIKETA_is3800-InspectionID" <> #Kamera.last_id_etiketa THEN
               #Kamera.last_id_etiketa := "COG_ETIKETA_is3800-InspectionID";
               IF #Kamera.sber_aktivni THEN
                   #Kamera.prijato_etiketa := TRUE;
               END_IF;
           END_IF;
           // text prevzit, jakmile je k dispozici (i o par cyklu pozdeji nez ID);
           // prazdny vysledek dalsi inspekce dobry text neprepise
           IF #Kamera.sber_aktivni AND #Kamera.prijato_etiketa AND "DB_data_ctena".upraveny <> '' THEN
               #Kamera.text_etiketa := "DB_data_ctena".upraveny;
               #Kamera.ok_etiketa := TRUE;
           END_IF;
           IF "COG_FOLIE_L_is3800-InspectionID" <> #Kamera.last_id_folie_l THEN
               #Kamera.last_id_folie_l := "COG_FOLIE_L_is3800-InspectionID";
               IF #Kamera.sber_aktivni THEN
                   #Kamera.prijato_folie_l := TRUE;
                   #Kamera.ok_folie_l := ("COG_FOLIE_L_is3800-InspectionResults[0]" OR "COG_FOLIE_L_is3800-InspectionResults[1]") <> 16#00;
               END_IF;
           END_IF;
           IF "COG_FOLIE_P_is3800-InspectionID" <> #Kamera.last_id_folie_p THEN
               #Kamera.last_id_folie_p := "COG_FOLIE_P_is3800-InspectionID";
               IF #Kamera.sber_aktivni THEN
                   #Kamera.prijato_folie_p := TRUE;
                   #Kamera.ok_folie_p := ("COG_FOLIE_P_is3800-InspectionResults[0]" OR "COG_FOLIE_P_is3800-InspectionResults[1]") <> 16#00;
               END_IF;
           END_IF;
       END_REGION

       REGION Timeout - plato opustilo s2 a vysledky nedorazily
           #TIMER.TIMER_6.TON(IN := #Kamera.sber_aktivni AND NOT #SENSORS.kontrola,
                              PT := #Kamera.timeout_sberu);
       END_REGION

       REGION Vyhodnoceni a zapis do fronty
           IF #Kamera.sber_aktivni AND
               ((#Kamera.prijato_etiketa AND #Kamera.prijato_folie_l AND #Kamera.prijato_folie_p)
               OR #TIMER.TIMER_6.Q OR #Kamera.s2_nabeh) THEN

               #ocekavany_text := CONCAT(IN1 := "DB_HMI_recype".recipe.pole_string_2,
                                         IN2 := "DB_HMI_recype".recipe.pole_string_1);
               #format_etiketa_ok := #Kamera.bypass_ocr
               OR (FIND(IN1 := #Kamera.text_etiketa, IN2 := "DB_HMI_recype".recipe.pole_string_2) > 0
               AND NOT "OP2_DB".Tisk.datum_chyba);

               // kontrola kodu tridirny - nezavisla na bypass_ocr, vypinatelna z HMI
               #Kamera.tridirna_ok := NOT #Kamera.kontrola_tridirny
               OR FIND(IN1 := #Kamera.text_etiketa, IN2 := #KOD_TRIDIRNY) > 0;

               #Kamera.vyradit := NOT #Kamera.prijato_etiketa OR NOT #Kamera.prijato_folie_l
               OR NOT #Kamera.prijato_folie_p OR NOT #Kamera.ok_etiketa
               OR NOT #format_etiketa_ok OR NOT #Kamera.ok_folie_l
               OR NOT #Kamera.ok_folie_p
               OR NOT #Kamera.tridirna_ok;

               IF #Kamera.text_etiketa = '' THEN
                   #Kamera.text_etiketa := 'NECTENO';   // prazdny text = prazdna pozice!
               END_IF;

               // zapis ZA posledni obsazenou pozici
               #Kamera.idx := 0;
               FOR #i := 5 TO 1 BY -1 DO
                   IF "DB_HMI_recype".fronta[#i].prenaseny_text <> '' THEN
                       #Kamera.idx := #i;
                       EXIT;
                   END_IF;
               END_FOR;

               IF #Kamera.idx < 5 THEN
                   "DB_HMI_recype".fronta[#Kamera.idx + 1].prenaseny_text := #Kamera.text_etiketa;
                   "DB_HMI_recype".fronta[#Kamera.idx + 1].balik_den := #Kamera.balik_den;
                   "DB_HMI_recype".fronta[#Kamera.idx + 1].vyrazeni := #Kamera.vyradit;
               ELSE
                   #Kamera.fronta_plna := TRUE;
               END_IF;
               #Kamera.sber_aktivni := FALSE;
           END_IF;
       END_REGION

       REGION Novy balik pod kamerou - start sberu (az PO zapisu predchoziho)
           IF #Kamera.s2_nabeh THEN
               // citac plat (presunuto ze site 20)
               #zpracovani_dat[1].balik_den := #zpracovani_dat[1].balik_den + 1;
               IF #zpracovani_dat[1].balik_den >= 32000 THEN
                   #zpracovani_dat[1].balik_den := 1;
               END_IF;
               #Kamera.balik_den := #zpracovani_dat[1].balik_den;   // az PO pricteni

               #Kamera.sber_aktivni := TRUE;
               #Kamera.prijato_etiketa := FALSE;
               #Kamera.prijato_folie_l := FALSE;
               #Kamera.prijato_folie_p := FALSE;
               #Kamera.ok_etiketa := FALSE;
               #Kamera.ok_folie_l := FALSE;
               #Kamera.ok_folie_p := FALSE;
               #Kamera.text_etiketa := '';
           END_IF;
       END_REGION
   END_IF;

   REGION Obsazenost fronty pro HMI (pocita se kazdy scan)
       #Kamera.pocet := 0;
       FOR #i := 1 TO 5 DO
           IF "DB_HMI_recype".fronta[#i].prenaseny_text <> '' THEN
               #Kamera.pocet := #Kamera.pocet + 1;
           END_IF;
       END_FOR;
       "DB_HMI_recype".obsazenost_fronty := #Kamera.pocet;
       IF #Kamera.pocet = 0 THEN
           #Kamera.fronta_plna := FALSE;
       END_IF;
   END_REGION
END_REGION

REGION Network 22 (SCL): PŘEPNUTÍ JOBU HORNÍ KAMERY
   // Prepnuti jobu horni kamery podle receptury.
   // Spousti se nabeznou hranou "DB_HMI_recype".ODESLI_dATA (tlacitko Odeslani dat do tiskarny)
   // - soubezne s odeslanim zpravy do tiskarny (OP2).
   // Job 0 v recepture = job neprepinat.

   #Kam_Etiketa_Job.pozadovany := "DB_HMI_recype".recipe.PRG_CAM_etiketa;

   IF "CONTROL_LINE_DB".trig.reset_error_all THEN
       #Kam_Etiketa_Job.chyba := FALSE;
   END_IF;

   CASE #Kam_Etiketa_Job.krok OF
       0:  // ---- klid: cekam na pozadavek ----
           #Kam_Etiketa_Job.aktivni := FALSE;
           "COG_ETIKETA_is3800-ExecuteCommand/JobLoad" := FALSE;
           IF "DB_HMI_recype".ODESLI_dATA AND NOT #Kam_Etiketa_Job.odesli_pamet
               AND #Kam_Etiketa_Job.pozadovany > 0
               AND "COG_ETIKETA_is3800-Online" THEN
               "COG_ETIKETA_is3800-CommandID" := INT_TO_WORD(#Kam_Etiketa_Job.pozadovany);
               #Kam_Etiketa_Job.aktivni := TRUE;
               #Kam_Etiketa_Job.chyba := FALSE;
               #Kam_Etiketa_Job.krok := 10;
           END_IF;

       10: // ---- CommandID uz je venku (predchozi cyklus) -> spustit prikaz ----
           "COG_ETIKETA_is3800-ExecuteCommand/JobLoad" := TRUE;
           #Kam_Etiketa_Job.krok := 20;

       20: // ---- cekam na vysledek ----
           IF "COG_ETIKETA_is3800-CommandCompleted" THEN
               #Kam_Etiketa_Job.krok := 30;
           ELSIF "COG_ETIKETA_is3800-CommandFailed" THEN
               #Kam_Etiketa_Job.chyba := TRUE;
               #Kam_Etiketa_Job.chyba_kod := "COG_ETIKETA_is3800-CommandResultCode";
               #Kam_Etiketa_Job.krok := 30;
           ELSIF #TIMER.TIMER_3.Q THEN
               #Kam_Etiketa_Job.chyba := TRUE;            // kamera neodpovedela
               #Kam_Etiketa_Job.chyba_kod := 16#FFFF;
               #Kam_Etiketa_Job.krok := 30;
           END_IF;

       30: // ---- ukonceni handshake: shodit Execute, pockat az kamera shodi stav ----
           "COG_ETIKETA_is3800-ExecuteCommand/JobLoad" := FALSE;
           IF NOT "COG_ETIKETA_is3800-CommandCompleted"
               AND NOT "COG_ETIKETA_is3800-CommandFailed" THEN
               #Kam_Etiketa_Job.krok := 0;
           END_IF;

       ELSE
           #Kam_Etiketa_Job.krok := 0;
   END_CASE;

   // casovac timeoutu bezi v krocich 10..30
   #TIMER.TIMER_3.TON(IN := #Kam_Etiketa_Job.krok >= 10,
                      PT := #Kam_Etiketa_Job.timeout);
   IF #TIMER.TIMER_3.Q AND #Kam_Etiketa_Job.krok = 30 THEN
       #Kam_Etiketa_Job.krok := 0;                         // pojistka, kdyby kamera stav neshodila
   END_IF;

   #Kam_Etiketa_Job.odesli_pamet := "DB_HMI_recype".ODESLI_dATA;

   // kontrola: v klidu musi job v kamere odpovidat recepture
   #Kam_Etiketa_Job.nesouhlasi := #Kam_Etiketa_Job.krok = 0
   AND #Kam_Etiketa_Job.pozadovany > 0
   AND "COG_ETIKETA_is3800-Online"
   AND WORD_TO_INT("COG_ETIKETA_is3800-Current Job ID") <> #Kam_Etiketa_Job.pozadovany;
END_REGION

REGION Network 23: EXTERNAL_TRIGER
   RUNG wire#powerrail
      { S7_Templates := "SrcType := Int" } EQ_Contact(in1 := #SQCR, in2 := #STEP_5_HOME)
      Contact( "INICIALIZACE_RUN" )
      I_Contact( #TRIG.inicial_ok_op )
      Contact( "AUTOMAT" )
      S_Coil( #HMI.reset_fronty )
      S_Coil( #TRIG.inicial_ok_op )
   END_RUNG
   RUNG wire#powerrail
      Contact( "FirstScan" )
      S_Coil( #HMI.reset_fronty )
      Move(in := 0, out1 => "DB_HMI_recype".obsazenost_fronty, out2 => #zpracovani_dat[1].balik_den)
   END_RUNG
   // the same network as SCL:
   IF (#SQCR = #STEP_5_HOME) AND "INICIALIZACE_RUN" AND NOT #TRIG.inicial_ok_op AND "AUTOMAT" THEN
       #HMI.reset_fronty := TRUE;
       #TRIG.inicial_ok_op := TRUE;
   END_IF;
   IF "FirstScan" THEN
       #HMI.reset_fronty := TRUE;
       "DB_HMI_recype".obsazenost_fronty := 0;
       #zpracovani_dat[1].balik_den := 0;
   END_IF;
END_REGION

REGION Network 24: ETERNAL_TRIGR_INICIAL
   RUNG wire#powerrail
      Contact( "AUTOMAT" )
      { S7_Templates := "SrcType := Int" } GT_Contact(in1 := #SQCR, in2 := #STEP_0)
      { S7_Templates := "SrcType := Int" } LT_Contact(in1 := #SQCR, in2 := #STEP_1000)
      I_Contact( #Kam_Etiketa_Job.aktivni )
      Coil( "COG_ETIKETA_COG_ETIKETA_is3800-TriggerEnable" )
   END_RUNG
   RUNG wire#powerrail
      Contact( "AUTOMAT" )
      { S7_Templates := "SrcType := Int" } GT_Contact(in1 := #SQCR, in2 := #STEP_0)
      { S7_Templates := "SrcType := Int" } LT_Contact(in1 := #SQCR, in2 := #STEP_1000)
      Coil( "COG_FOLIE_L_COG_FOLIE_L_is3800-TriggerEnable" )
   END_RUNG
   RUNG wire#powerrail
      Contact( "AUTOMAT" )
      { S7_Templates := "SrcType := Int" } GT_Contact(in1 := #SQCR, in2 := #STEP_0)
      { S7_Templates := "SrcType := Int" } LT_Contact(in1 := #SQCR, in2 := #STEP_1000)
      Coil( "COG_FOLIE_P_COG_FOLIE_P_is3800-TriggerEnable" )
   END_RUNG
   // the same network as SCL:
   "COG_ETIKETA_COG_ETIKETA_is3800-TriggerEnable" := "AUTOMAT" AND (#SQCR > #STEP_0) AND (#SQCR < #STEP_1000) AND NOT #Kam_Etiketa_Job.aktivni;
   "COG_FOLIE_L_COG_FOLIE_L_is3800-TriggerEnable" := "AUTOMAT" AND (#SQCR > #STEP_0) AND (#SQCR < #STEP_1000);
   "COG_FOLIE_P_COG_FOLIE_P_is3800-TriggerEnable" := "AUTOMAT" AND (#SQCR > #STEP_0) AND (#SQCR < #STEP_1000);
END_REGION

REGION Network 25: hmi
END_REGION

REGION Network 26 (SCL): VYRAZENI MANUAL
   (* #Test_tp_ka12(IN := "DB_Manual".test_vyr,
                 PT := T#500MS);

   "-KA12" := #Test_tp_ka12.Q;

   // testovací bit se sám shodí → každý Modify TRUE = jeden pulz
   IF "DB_Manual".test_vyr THEN
       "DB_Manual".test_vyr := FALSE;
   END_IF; *)
END_REGION
END_FUNCTION_BLOCK
